Staubli VAL3: isDefine.pgx

public program isDefine(string x_sKey, bool& x_bResult)
begin
  x_bResult=isDefined(trajTemp:tTrajItem[x_sKey])
end
